(* IEC 61131-3 sources: axsharp/src/AXSharp.compiler/tests/integration/expected/app/src, 2 files *)

(* ---- configuration.st ---- *)
CONFIGURATION MyConfiguration
    TASK Main(Interval := T#1000ms, Priority := 1);
    PROGRAM P1 WITH Main: MyProgram;

    VAR_GLOBAL
	{S7.extern=ReadWrite}
        lib1_MyClass : lib1.MyClass;
	{S7.extern=ReadWrite}
        lib2_MyClass : lib2.MyClass;
    END_VAR
END_CONFIGURATION

(* ---- program.st ---- *)
PROGRAM MyProgram
    VAR_EXTERNAL

    END_VAR

    VAR

    END_VAR

    VAR_TEMP

    END_VAR

    // code here
    ;
END_PROGRAM
